(* IEC 61131-3 sources: plc-hackathon-2026/work/dump/MyController/Plc Logic/Application/Date_and_Time, 3 files *)

(* ---- GVL_HMI.st ---- *)
VAR_GLOBAL
	// PLC datum i vrijeme - DT format SET
	PLC_Datum_Vrijeme_Get_DT : DT;
	// PLC datum i vrijeme - trenutna godina
	PLC_Datum_Vrijeme_Godina AT %MW490: INT;
	// PLC datum i vrijeme - trenutni mjesec
	PLC_Datum_Vrijeme_Mjesec AT %MW491: INT;
	// PLC datum i vrijeme - trenutni dan
	PLC_Datum_Vrijeme_Dan AT %MW492: INT;
	// PLC datum i vrijeme - trenutni sat
	PLC_Datum_Vrijeme_Sat AT %MW493: INT;
	// PLC datum i vrijeme - trenutna minuta
	PLC_Datum_Vrijeme_Minuta AT %MW494: INT;
	// PLC datum i vrijeme - trenutna sekunda
	PLC_Datum_Vrijeme_Sekunda AT %MW495: INT;

	// PLC datum i vrijeme - DT format GET
	PLC_Datum_Vrijeme_Set_DT : DT;
	promjeni : BOOL;

	// Parametar - PLC datum i vrijeme - godina
	PAR_PLC_Datum_Vrijeme_Godina AT %MW1020: INT;
	// Parametar - PLC datum i vrijeme - mjesec
	PAR_PLC_Datum_Vrijeme_Mjesec AT %MW1021: INT;
	// Parametar - PLC datum i vrijeme - dan
	PAR_PLC_Datum_Vrijeme_Dan AT %MW1022: INT;
	// Parametar - PLC datum i vrijeme - sat
	PAR_PLC_Datum_Vrijeme_Sat AT %MW1023: INT;
	// Parametar - PLC datum i vrijeme - minuta
	PAR_PLC_Datum_Vrijeme_Minuta AT %MW1024: INT;
	// Parametar - PLC datum i vrijeme - sekunda
	PAR_PLC_Datum_Vrijeme_Sekunda AT %MW1025: INT;
END_VAR

(* ---- Datum_Vrijeme_Get.st ---- *)
FUNCTION_BLOCK Datum_Vrijeme_Get
VAR_OUTPUT
	OUT_Date_Time : DT;
	OUT_Year : INT;
	OUT_Month : INT;
	OUT_Day : INT;
	OUT_Hour : INT;
	OUT_Minute : INT;
	OUT_Second : INT;
END_VAR
VAR
    uidResultRtcGet: UDINT;
	dwRtcGet: DWORD;
    stGetDate: SysTimeRtc.RTS_SYSTIMEDATE;
	udiGetSysTimeDate: RTS_IEC_RESULT;
    uiGetYear: UINT;
    uiGetMonth: UINT;
    uiGetDay: UINT;
    uiGetHour: UINT;
    uiGetMinute: UINT;
    uiGetSecond: UINT;
    uiGetMSecond: UINT;
    uiGetDayOfWeek: UINT;
    uiGetYday: UINT;
    uidResultConvertToDate: UDINT;

	udiResultConvertToUtc: UDINT;
    stSetDate: SysTimeRtc.RTS_SYSTIMEDATE;
    dwSetTimeStamp: DWORD;
    xCommandSetRtc: BOOL;
    uidResultRtcSet: UDINT;

	Sekunda: BOOL;
	R_TRIG_Sekunda: R_TRIG;
	Always_Off: BOOL;
END_VAR

(* ---- Datum_Vrijeme_Set.st ---- *)
FUNCTION_BLOCK Datum_Vrijeme_Set
VAR_INPUT
	IN_Year : INT;
	IN_Month : INT;
	IN_Day : INT;
	IN_Hour : INT;
	IN_Minute : INT;
	IN_Second : INT;
END_VAR
VAR_OUTPUT
	OUT_Date_Time : DT;
END_VAR
VAR
    uidResultRtcGet: UDINT;
	dwRtcGet: DWORD;
    stGetDate: SysTimeRtc.RTS_SYSTIMEDATE;
	udiGetSysTimeDate: RTS_IEC_RESULT;
    uiGetYear: UINT;
    uiGetMonth: UINT;
    uiGetDay: UINT;
    uiGetHour: UINT;
    uiGetMinute: UINT;
    uiGetSecond: UINT;
    uiGetMSecond: UINT;
    uiGetDayOfWeek: UINT;
    uiGetYday: UINT;
    uidResultConvertToDate: UDINT;

	udiResultConvertToUtc: UDINT;
    stSetDate: SysTimeRtc.RTS_SYSTIMEDATE;
    dwSetTimeStamp: DWORD;
    xCommandSetRtc: BOOL;
    uidResultRtcSet: UDINT;

	Sekunda: BOOL;
	R_TRIG_Sekunda: R_TRIG;
	Always_Off: BOOL;
END_VAR
